TEXTLIST TextList_E_Line_Target
  0 = 'Drain'
  1 = 'Tank_A'
  2 = 'Tank_B'
  3 = 'CIP'
   = ''
END_TEXTLIST

(* stored: Version 1.1.0.1, ProductVersion 3.1.4024.12
   TextList TextList_E_Line_Target: Id {202b6309-6e0b-4fbc-9bc1-6fe68100ec53} *)
